TYPE ST_EL3xx4 :
STRUCT
	
	//4CH AI, RTD RES SNS
	State	AT %I*: UINT;

	ai_ch1	AT %I*: INT;
	ai_ch2	AT %I*: INT;
	ai_ch3	AT %I*: INT;
	ai_ch4	AT %I*: INT;
	
	
END_STRUCT
END_TYPE

(* stored: Version 1.1.0.1, ProductVersion 3.1.4024.12
   DUT ST_EL3xx4: Id {af02ebb4-0524-4452-b034-9a9500025db7} *)
